// POUs/_FB_ConfigXtsLoop
(****************************************************************************************************<br>
© Syntegon Group.<br>
All rights reserved, also regarding any disposal, exploitation, reproduction, editing, distribution,<br>
as well as in the event of applications for industrial property rights.<br>
*****************************************************************************************************<br>
DESCRIPTION:<br>
Parameter set of one XTS loop (ADR 0017): its pose, origin shift, track modules, zones and gripper fingers,<br>
written by the configurator, taken over when the application allows it. Typical cycle:<br>
  fb_FxxParam.m_Register(vio_Manifest := GVL_Config.stManifest, vi_udn_Id := fb_Fxx.m_Id());<br>
  fb_FxxParam.m_Cycle(vio_Default := FxxDefault, vio_Set := FxxSet, vi_b_ApplyAllowed := b_Stopped);<br>
  fb_Fxx.m_Configure(vi_Pose := fb_FxxParam.m_Pose(), vi_lr_ToolOffset := 120, ...);<br>
  fb_FxxParam.m_PassOn(vio_Visu := fb_Fxx);<br>
The application's logic takes its track and zones from m_Active, not from its own constants.<br>
*****************************************************************************************************<br>
OUTPUT VALUES:<br>
vo_Config is the contract structure the gateway reads and writes at the path in the config manifest.<br>
*****************************************************************************************************<br>
VERSION         ¦ DATE       ¦ NAME      ¦ CHANGE<br>
Syn_Config 1.1.0 ¦ 2026-11-10 ¦ J.Willner ¦ New<br>
Syn_Config 2.0.0 ¦ 2026-11-11 ¦ J.Willner ¦ Gripper fingers with their offsets (ADR 0018)<br>
****************************************************************************************************)
FUNCTION_BLOCK _FB_ConfigXtsLoop EXTENDS _FB_ConfigComponent
VAR_OUTPUT
	vo_Config							: ST_ConfigXtsLoop;	// contract structure of the gateway
END_VAR

(****************************************************************************************************<br>
© Syntegon Group.<br>
All rights reserved, also regarding any disposal, exploitation, reproduction, editing, distribution,<br>
as well as in the event of applications for industrial property rights.<br>
*****************************************************************************************************<br>
DESCRIPTION:<br>
All effective values (track modules, zones, ...), for the application's own logic.<br>
****************************************************************************************************)
METHOD m_Active : ST_ConfigXtsLoopParam
m_Active := vo_Config.stActive;
END_METHOD

(****************************************************************************************************<br>
© Syntegon Group.<br>
All rights reserved, also regarding any disposal, exploitation, reproduction, editing, distribution,<br>
as well as in the event of applications for industrial property rights.<br>
*****************************************************************************************************<br>
DESCRIPTION:<br>
An XTS loop.<br>
****************************************************************************************************)
METHOD PROTECTED m_ComponentType : SynVisu.E_VisuComponentType
m_ComponentType := SynVisu.E_VisuComponentType.XTS_LOOP;
END_METHOD

(****************************************************************************************************<br>
© Syntegon Group.<br>
All rights reserved, also regarding any disposal, exploitation, reproduction, editing, distribution,<br>
as well as in the event of applications for industrial property rights.<br>
*****************************************************************************************************<br>
DESCRIPTION:<br>
Every cycle: handles a staged set or a reset (a set only while vi_b_ApplyAllowed), keeps the active set in<br>
vio_Set and gives the effective values in vo_Config.stActive: the active set while one is valid, else the<br>
program values vio_Default.<br>
*****************************************************************************************************<br>
OUTPUT VALUES:<br>
TRUE in the cycle a set was taken over or reset.<br>
****************************************************************************************************)
METHOD m_Cycle : BOOL
VAR_IN_OUT CONSTANT
	vio_Default							: ST_ConfigXtsLoopParam;	// the application's program values
END_VAR
VAR_IN_OUT
	vio_Set								: ST_ConfigXtsLoopSet;	// the application's VAR PERSISTENT active set
END_VAR
VAR_INPUT
	vi_b_ApplyAllowed					: BOOL;	// [-] a staged set may be taken over now, e.g. while the machine stands
END_VAR
VAR
	str_TempRejection					: STRING(80);
END_VAR
m_Cycle := FALSE;
CASE m_Staging(vio_Staging := vo_Config.stStaging, vio_Status := vo_Config.stStatus, vi_b_ApplyAllowed := vi_b_ApplyAllowed,
	vi_udn_ActiveVersion := SEL(vio_Set.bValid, 0, vio_Set.nVersion)) OF
	E_ConfigAction.RESET:
		vio_Set.bValid := FALSE;
		m_Handled(vio_Staging := vo_Config.stStaging, vio_Status := vo_Config.stStatus, vi_str_Rejection := '');
		m_Cycle := TRUE;
	E_ConfigAction.TAKE_OVER:
		str_TempRejection := m_Invalid(vio_Param := vo_Config.stStaged);
		IF str_TempRejection = '' THEN
			vio_Set.nLastVersion := vio_Set.nLastVersion + 1;
			vio_Set.nVersion := vio_Set.nLastVersion;
			vio_Set.stParam := vo_Config.stStaged;
			vio_Set.bValid := TRUE;
			m_Cycle := TRUE;
		END_IF
		m_Handled(vio_Staging := vo_Config.stStaging, vio_Status := vo_Config.stStatus, vi_str_Rejection := str_TempRejection);
END_CASE


(****************************************************************************************************
EFFECTIVE VALUES
****************************************************************************************************)
IF vio_Set.bValid THEN
	vo_Config.stActive := vio_Set.stParam;
	vo_Config.stStatus.nActiveVersion := vio_Set.nVersion;
ELSE
	vo_Config.stActive := vio_Default;
	vo_Config.stStatus.nActiveVersion := 0;
END_IF
END_METHOD

(****************************************************************************************************<br>
© Syntegon Group.<br>
All rights reserved, also regarding any disposal, exploitation, reproduction, editing, distribution,<br>
as well as in the event of applications for industrial property rights.<br>
*****************************************************************************************************<br>
DESCRIPTION:<br>
Why a staged set cannot be taken over; '' when it can: a track without modules, more modules, zones or fingers<br>
than the lists hold, a module without a length, a zone on no conveyor (id 0), or a finger without a diameter or<br>
height.<br>
****************************************************************************************************)
METHOD PRIVATE m_Invalid : STRING(80)
VAR_IN_OUT CONSTANT
	vio_Param							: ST_ConfigXtsLoopParam;	// the staged set
END_VAR
m_Invalid := m_InvalidModules(vio_aModules := vio_Param.aModules, vi_un_Count := vio_Param.nModuleCount);
IF m_Invalid = '' THEN
	m_Invalid := m_InvalidZones(vio_aZones := vio_Param.aZones, vi_un_Count := vio_Param.nZoneCount);
END_IF
IF m_Invalid = '' THEN
	m_Invalid := m_InvalidFingers(vio_aFingers := vio_Param.aFingers, vi_un_Count := vio_Param.nFingerCount);
END_IF
END_METHOD

(****************************************************************************************************<br>
© Syntegon Group.<br>
All rights reserved, also regarding any disposal, exploitation, reproduction, editing, distribution,<br>
as well as in the event of applications for industrial property rights.<br>
*****************************************************************************************************<br>
DESCRIPTION:<br>
Passes the effective origin shift, track modules, zones and fingers on to the loop's Syn_Visu FB, so the<br>
visualisation shows what the machine uses. The pose goes with the application's own m_Configure call (with<br>
the tool offset and mover size, hardware): vi_Pose := m_Pose(). Call it after m_Cycle, every cycle; Syn_Visu's<br>
config version only changes when a value does.<br>
****************************************************************************************************)
METHOD m_PassOn : BOOL
VAR_IN_OUT
	vio_Visu							: SynVisu._FB_VisuXtsLoop;	// the loop's Syn_Visu FB
END_VAR
m_PassOn := TRUE;
vio_Visu.m_SetOriginShift(vi_lr_X := vo_Config.stActive.stOriginShift.fX, vi_lr_Y := vo_Config.stActive.stOriginShift.fY,
	vi_lr_Z := vo_Config.stActive.stOriginShift.fZ);
m_PassOnModules(vio_Visu := vio_Visu, vio_aModules := vo_Config.stActive.aModules,
	vi_un_Count := vo_Config.stActive.nModuleCount, vi_un_VisuCount := vio_Visu.vo_Visu.stConfig.nModuleCount);
m_PassOnZones(vio_Visu := vio_Visu, vio_aZones := vo_Config.stActive.aZones, vi_un_Count := vo_Config.stActive.nZoneCount,
	vi_un_VisuCount := vio_Visu.vo_Visu.stConfig.nZoneCount);
m_PassOnFingers(vio_Visu := vio_Visu, vio_aFingers := vo_Config.stActive.aFingers,
	vi_un_Count := vo_Config.stActive.nFingerCount, vi_un_VisuCount := vio_Visu.vo_Visu.stConfig.nFingerCount);
END_METHOD

(****************************************************************************************************<br>
© Syntegon Group.<br>
All rights reserved, also regarding any disposal, exploitation, reproduction, editing, distribution,<br>
as well as in the event of applications for industrial property rights.<br>
*****************************************************************************************************<br>
DESCRIPTION:<br>
Effective pose of the start of module 1 (MCS), for the application's logic and its Syn_Visu m_Configure call.<br>
****************************************************************************************************)
METHOD m_Pose : SynVisu.ST_VisuPose
m_Pose := vo_Config.stActive.stPose;
END_METHOD

END_FUNCTION_BLOCK

// POUs/_FC_GetVersionSynConfig
(****************************************************************************************************<br>
© Syntegon Group.<br>
All rights reserved, also regarding any disposal, exploitation, reproduction, editing, distribution,<br>
as well as in the event of applications for industrial property rights.<br>
*****************************************************************************************************<br>
DESCRIPTION:<br>
Runtime-readable version of the Syn_Config library.<br>
*****************************************************************************************************<br>
VERSION         ¦ DATE       ¦ NAME      ¦ CHANGE<br>
Syn_Config 1.0.0 ¦ 2026-11-10 ¦ J.Willner ¦ Parameter sets of conveyors and Deltas (ADR 0017, protocol 1)<br>
Syn_Config 1.1.0 ¦ 2026-11-10 ¦ J.Willner ¦ Every other component type (#24)<br>
Syn_Config 2.0.0 ¦ 2026-11-11 ¦ J.Willner ¦ Gripper fingers in the robots' sets (protocol 2, #25)<br>
****************************************************************************************************)
FUNCTION _FC_GetVersionSynConfig : UINT
VAR_INPUT
	vi_n_VersionElement					: INT;	// [-] 1 = major, 2 = minor, 3 = revision
END_VAR

CASE vi_n_VersionElement OF
	1: _FC_GetVersionSynConfig := 2;
	2: _FC_GetVersionSynConfig := 0;
	3: _FC_GetVersionSynConfig := 0;
ELSE
	_FC_GetVersionSynConfig := 16#FFFF;
END_CASE

END_FUNCTION
